FUNCTION_BLOCK Heat_Control_Slider (* Composite Function Block Type *)
  (* Standard: 61499-2 *)
  (* Version 0.0, 12/30/2019, prana, nxtControl GmbH, template *)
  PACKAGE Main;
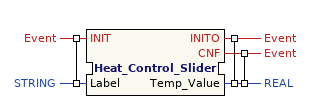
  EVENT_INPUT
    INIT WITH Label; (* Initialization Request *)
  END_EVENT
  EVENT_OUTPUT
    INITO WITH Temp_Value; (* Initialization Confirm *)
    CNF WITH Temp_Value; (* Execution Confirmation *)
  END_EVENT
  VAR_INPUT
    Label : STRING; (* Input event qualifier *)
  END_VAR
  VAR_OUTPUT
    Temp_Value : REAL := 40; (* Output event qualifier *)
  END_VAR
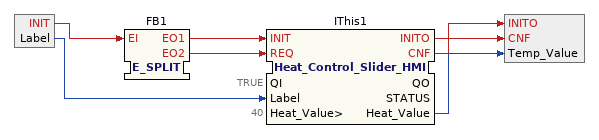
  FBS
    IThis1 : Heat_Control_Slider_HMI(Heat_Value> := 40, QI := TRUE);
    FB1 : E_SPLIT;
  END_FBS
  EVENT_CONNECTIONS
    INIT TO FB1.EI;
    FB1.EO1 TO IThis1.INIT;
    FB1.EO2 TO IThis1.REQ;
    IThis1.INITO TO INITO;
    IThis1.CNF TO CNF;
  END_CONNECTIONS
  DATA_CONNECTIONS
    Label TO IThis1.Label;
    IThis1.Heat_Value TO Temp_Value;
  END_CONNECTIONS
END_FUNCTION_BLOCK
